RoboDK station: hand_motion.rdk

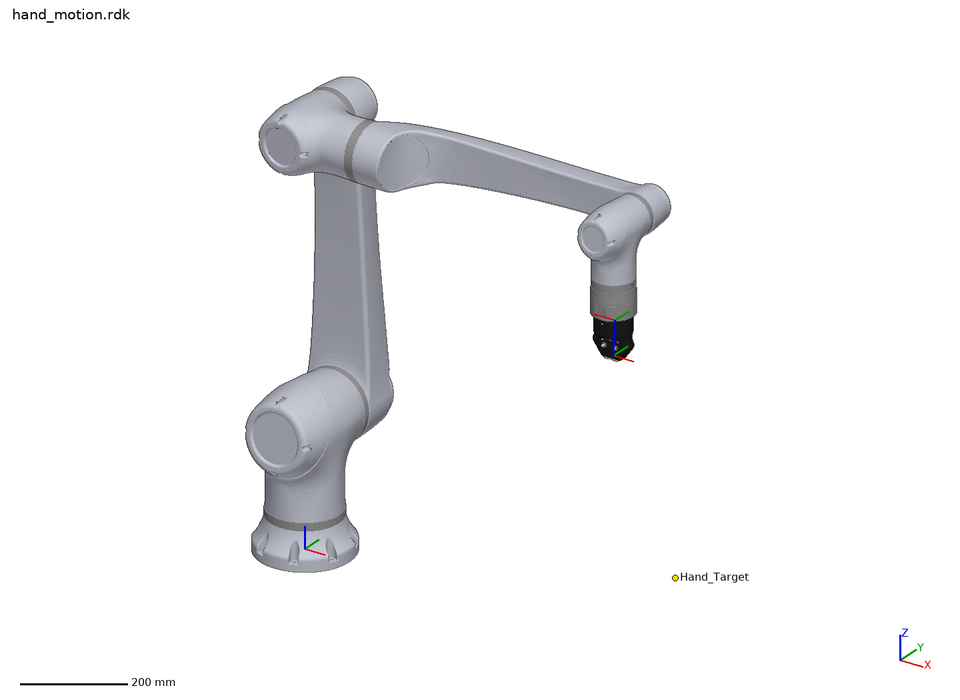
[picture v0: the station drawn from its stored meshes, robots at their saved joint values, targets as dots, program paths as lines]
Station hand_motion (saved by RoboDK 6.0.3). Poses are relative to the parent item; angles as X-Y-Z fixed-axis rotations.
  - frame Neura LARA 8 Base at (0, 0, 0) mm
    - robot Neura LARA 8: 6 axes
        modified DH rows (alpha deg, a mm, theta deg, d mm): 0, 0, 0, 260; -90, 0, -90, 0; 0, 600, -90, 0; -90, 0, 0, 700; 90, 0, 0, 0; -90, 0, 180, 179.5
        joint limits [-180, -135, -155, -180, -180, -360] to [180, 135, 155, 180, 180, 360]; home [0, 0, 90, 0, 90, 0]; saved at [0, 0, 90, 0, 90, 0]
      - robot RobotiQ 2F-85 Gripper (Mechanism) (model RobotiQ 2F85): 1 axes, payload 5 kg
          joint limits [0] to [85]; home [85]; saved at [0]
        - frame Grip_Attach_Frame at (-4.53, -1.14, 10.96) mm
    - target Hand_Target (Cartesian target) at (819.81, 29.81, 156.61) mm, rotated rx 180 ry 0 rz -180 deg; joints [4.563, 26.506, 87.684, 0, 65.81, 4.563] of Neura LARA 8
  - object Cube 50mm at (805.02, 3.79, 48.01) mm, rotated rx 180 ry 0 rz -174.82 deg, size 50 x 50 x 50 mm, geometry from Cube-50mm.sld
  - frame RobotiQ 2F-85 Gripper (Mechanism) Base at (0, 1000, 0) mm
